PROGRAM POU
VAR
	FB_ValveControl_0: FB_ValveControl;
	Actual_ValveMode: BYTE;
	
	SetValaveMode: BYTE;
	SetAppControl: BYTE;
	SetAppOption: BYTE;
	SetpointValue1: INT;
	SetpointValue2: INT;
	Acknowledge: BOOL;
	ActualValveState: BYTE;
	ActualAppState: BYTE;
	ActualValue1: INT;
	ActualValue2: INT;
	Response: eResponseToValveModeSet;
	ErrorCode: INT;
	FB_Upload_Single_Parameter_0: FB_Upload_Single_Parameter;
	Upload_Execute: BOOL;
	Upload_Channel: INT;
	Upld_AddrTarget: INT;
	Upload_Index: INT;
	Upld_Response: Festo_VTEM.eTransferResponse;
	Uploaded_Value: INT;
	Upload_Done: BOOL;
	Upload_Error: BOOL;
	FB_Download_Single_Parameter_0: FB_Download_Single_Parameter;
	Download_Execute: BOOL;
	Download_Channel: INT;
	Dwnlad_AddrTarget: INT;
	Download_Index: INT;
	DownloadValue: INT;
	Download_Done: BOOL;
	Download_Error: BOOL;
	Dwnlad_Response: Festo_VTEM.eTransferResponse;
	FB_ReadMalfunctionList_0: FB_ReadMalfunctionList;
	Malf_Execute: BOOL;
	xAbort: BOOL;
	ChooseValve: USINT;
	Malf_List: ARRAY [1..40] OF Festo_VTEM.stMalfunction;
	Malfunction_Tiemstap: stTimeStamp;
	Malfunction_Response: eResponseReadMalfunctionList;
	Malfunction_Busy: BOOL;
	Malfunction_Done: BOOL;
	Malfunction_Error: BOOL;
	Malfunction_Aborted: BOOL;
	FB_Save_Configuration_Persistent_0: FB_Save_Configuration_Persistent;
	Save_Execute: BOOL;
	Save_Done: BOOL;
	Save_Error: BOOL;
	Save_Response: Festo_VTEM.eSavingResponse;
	Enable: BOOL;
END_VAR

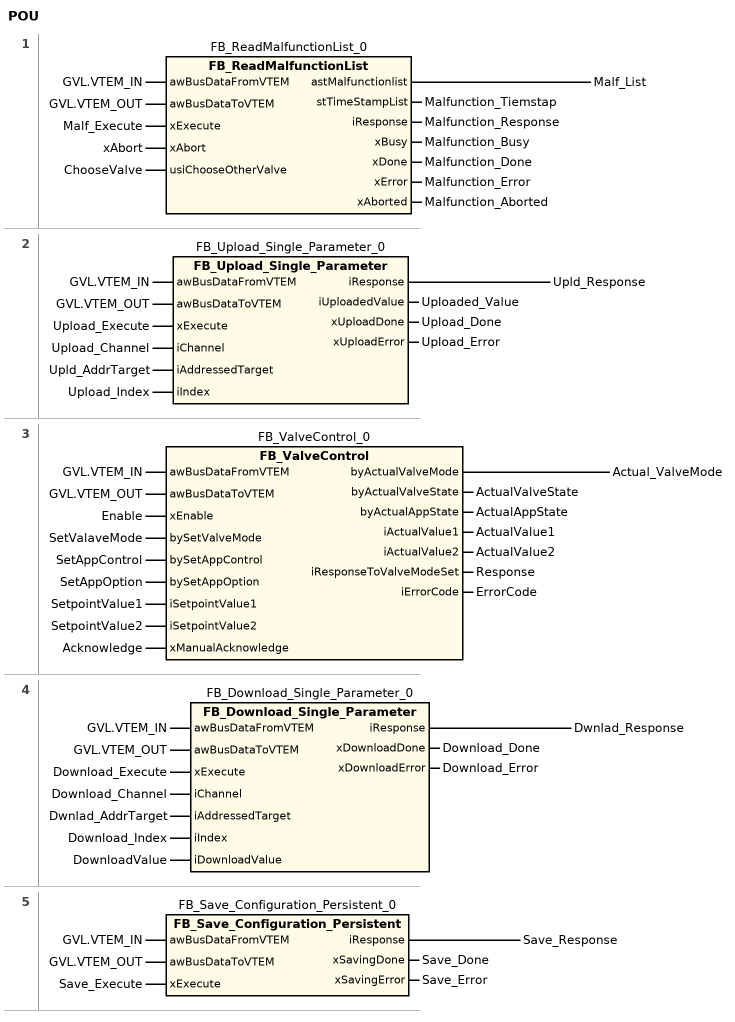
// NETWORK 1
FB_ReadMalfunctionList_0(
    awBusDataFromVTEM := GVL.VTEM_IN,
    awBusDataToVTEM := GVL.VTEM_OUT,
    xExecute := Malf_Execute,
    xAbort := xAbort,
    usiChooseOtherValve := ChooseValve,
    stTimeStampList => Malfunction_Tiemstap,
    iResponse => Malfunction_Response,
    xBusy => Malfunction_Busy,
    xDone => Malfunction_Done,
    xError => Malfunction_Error,
    xAborted => Malfunction_Aborted); // FB_ReadMalfunctionList
Malf_List := FB_ReadMalfunctionList_0.astMalfunctionlist;

// NETWORK 2
FB_Upload_Single_Parameter_0(
    awBusDataFromVTEM := GVL.VTEM_IN,
    awBusDataToVTEM := GVL.VTEM_OUT,
    xExecute := Upload_Execute,
    iChannel := Upload_Channel,
    iAddressedTarget := Upld_AddrTarget,
    iIndex := Upload_Index,
    iUploadedValue => Uploaded_Value,
    xUploadDone => Upload_Done,
    xUploadError => Upload_Error); // FB_Upload_Single_Parameter
Upld_Response := FB_Upload_Single_Parameter_0.iResponse;

// NETWORK 3
FB_ValveControl_0(
    awBusDataFromVTEM := GVL.VTEM_IN,
    awBusDataToVTEM := GVL.VTEM_OUT,
    xEnable := Enable,
    bySetValveMode := SetValaveMode,
    bySetAppControl := SetAppControl,
    bySetAppOption := SetAppOption,
    iSetpointValue1 := SetpointValue1,
    iSetpointValue2 := SetpointValue2,
    xManualAcknowledge := Acknowledge,
    byActualValveState => ActualValveState,
    byActualAppState => ActualAppState,
    iActualValue1 => ActualValue1,
    iActualValue2 => ActualValue2,
    iResponseToValveModeSet => Response,
    iErrorCode => ErrorCode); // FB_ValveControl
Actual_ValveMode := FB_ValveControl_0.byActualValveMode;

// NETWORK 4
FB_Download_Single_Parameter_0(
    awBusDataFromVTEM := GVL.VTEM_IN,
    awBusDataToVTEM := GVL.VTEM_OUT,
    xExecute := Download_Execute,
    iChannel := Download_Channel,
    iAddressedTarget := Dwnlad_AddrTarget,
    iIndex := Download_Index,
    iDownloadValue := DownloadValue,
    xDownloadDone => Download_Done,
    xDownloadError => Download_Error); // FB_Download_Single_Parameter
Dwnlad_Response := FB_Download_Single_Parameter_0.iResponse;

// NETWORK 5
FB_Save_Configuration_Persistent_0(
    awBusDataFromVTEM := GVL.VTEM_IN,
    awBusDataToVTEM := GVL.VTEM_OUT,
    xExecute := Save_Execute,
    xSavingDone => Save_Done,
    xSavingError => Save_Error); // FB_Save_Configuration_Persistent
Save_Response := FB_Save_Configuration_Persistent_0.iResponse;

END_PROGRAM

(* stored: Version 1.1.0.1, ProductVersion 3.1.4024.16
   POU POU: Id {a79124f9-a500-417b-868f-291cae013984}, SpecialFunc None *)
